// Position planaire (docs/05 § 6.1), toujours en frame 0
{attribute 'pack_mode' := '1'}
TYPE ST_PlanarPos :
STRUCT
    stPos : ST_Position;
    eKind : E_PlanarPosKind;
    nStation : USINT;
END_STRUCT
END_TYPE

(* stored: Version 1.1.0.1, ProductVersion 3.1.4024.12
   DUT ST_PlanarPos: Id {990e3ef1-263c-527f-a2ca-b1bd245f2994} *)
